(* IEC 61131-3 sources: codesys-to-s7/tests/corpus/C2S7-GFX-SFC/neg, 1 file *)

(* ---- input.st ---- *)
PROGRAM PRG_S
VAR
    i : INT;
END_VAR
i := i + 1;
END_PROGRAM
